// Bundles the services every catalog event needs (injected once).
INTERFACE I_EventContext

PROPERTY Texts : I_TextProvider
GET
END_GET
END_PROPERTY

PROPERTY Language : I_LanguageProvider
GET
END_GET
END_PROPERTY

PROPERTY Formatter : I_TextFormatter
GET
END_GET
END_PROPERTY

PROPERTY EventEntries : I_EventEntryProvider
GET
END_GET
END_PROPERTY

END_INTERFACE

(* stored: Version 1.1.0.1, ProductVersion 3.1.4026.26
   Itf I_EventContext: Id {0d591c57-3607-414a-8364-3eb5e085e64d}
   Property Texts: Id {4062910d-0f44-4210-a057-ae09ae161031}
   Get Get: Id {be4e4733-b8ed-404d-9d04-1fb8821344c5}
   Property Language: Id {bec90ce6-9602-4114-8eb5-8a121ab2b42e}
   Get Get: Id {f7dd4a45-af73-4d4f-be68-b8f66a302ca8}
   Property Formatter: Id {c95434e1-185f-4f97-aa53-d2f9e0a80257}
   Get Get: Id {a204f7b8-7205-48f0-b7c1-c44793f13b1e}
   Property EventEntries: Id {73f6f02c-cb9c-45a8-abaf-4a5a1d866f7c}
   Get Get: Id {87094983-449f-4589-81bc-1b9bd3d58fd4} *)
